TYPE ST_Gr05HMIRef :
STRUCT
	stHMITOPLC				:ST_Gr05HMITOPLC;
	stPLCTOHMI				:ST_Gr05PLCTOHMI;
END_STRUCT
END_TYPE

(* stored: Version 1.1.0.1, ProductVersion 3.1.4024.15
   DUT ST_Gr05HMIRef: Id {642180f9-6242-41ee-b425-cd7224361dbe} *)
